// TwinCAT 3 PLC project MainPLC
// ProgramVersion: 3.1.4026.20
// libraries:
//   Tc2_Standard, * (Beckhoff Automation GmbH)
//   Tc2_System, * (Beckhoff Automation GmbH)
// project tree:
//   DUTs/ stShutterCommand.TcDUT, eShutterCommandType.TcDUT, stShutterConfig.TcDUT, eShutterStateType.TcDUT, stShutterState.TcDUT, stSwitchConfig.TcDUT, eSwitchStateType.TcDUT, stSwitchState.TcDUT
//   GVLs/ gvlSwitches.TcGVL, gvlShutters.TcGVL
//   / PlcTask.TcTTO
//   POUs/ MAIN.TcPOU
//   POUs/Shutters/ fbShutter.TcPOU, fbShutterActuator.TcPOU, fbShutterController.TcPOU
//   POUs/Switches/ fbSwitch.TcPOU
// real-time tasks:
//   TASK PlcTask: cycle T#50000us, priority 20, ADS port 350
// I/O:
//   DEVICE Device 1 (EtherCAT), AmsNetId 169.254.52.30.2.1
//     Term 4 (EK1100) [EK1100 EtherCAT Coupler (2A E-Bus)]
//       Term 5 (EL1008) [EL1008 8Ch. Dig. Input 24V, 3ms]
//       Term 6 (EL1809) [EL1809 16Ch. Dig. Input 24V, 3ms]
//       Term 7 (EL1809) [EL1809 16Ch. Dig. Input 24V, 3ms]
//       Term 8 (EL1809) [EL1809 16Ch. Dig. Input 24V, 3ms]
//       Term 9 (EL1809) [EL1809 16Ch. Dig. Input 24V, 3ms]
//       Term 10 (EL1809) [EL1809 16Ch. Dig. Input 24V, 3ms]
//       Term 11 (EL2809) [EL2809 16Ch. Dig. Output 24V, 0.5A]
//       Term 12 (EL2809) [EL2809 16Ch. Dig. Output 24V, 0.5A]
//       Term 13 (EL2809) [EL2809 16Ch. Dig. Output 24V, 0.5A]
//       Term 14 (EL2809) [EL2809 16Ch. Dig. Output 24V, 0.5A]
//       Term 15 (EL9011) [EL9011 End Terminal]
// variable links:
//   MainPLC/MainPLC Instance <-> Device 1 (EtherCAT)/Term 4 (EK1100)/Term 11 (EL2809)
//     PlcTask Outputs/gvlShutters.gvShutter1Down <-> Channel 2/Output
//     PlcTask Outputs/gvlShutters.gvShutter1Up <-> Channel 1/Output
//   MainPLC/MainPLC Instance <-> Device 1 (EtherCAT)/Term 4 (EK1100)/Term 5 (EL1008)
//     PlcTask Inputs/gvlSwitches.gvSwitchR1Down <-> Channel 2/Input
//     PlcTask Inputs/gvlSwitches.gvSwitchR1Up <-> Channel 1/Input

CONFIGURATION MainPLC
    RESOURCE PLC ON TwinCAT3
        TASK PlcTask(INTERVAL := T#50000us, PRIORITY := 20);
        PROGRAM MAIN WITH PlcTask : MAIN;
    END_RESOURCE
END_CONFIGURATION

// ---- DUTs/stShutterCommand.TcDUT
TYPE stShutterCommand :
STRUCT
    CommandType  : eShutterCommandType;	// Command type
    Position : USINT;                	// Position for MOVE_TO_POSITION command
	Angle : USINT;						// Fin Angle for MOVE_TO_POSITION command
END_STRUCT
END_TYPE

// ---- DUTs/eShutterCommandType.TcDUT
{attribute 'qualified_only'}
{attribute 'strict'}
{attribute 'to_string'}
TYPE eShutterCommandType :
(
    NONE,           // No command
    OPEN,           // Open command (move to 100%)
    CLOSE,          // Close command (move to 0%)
	STEP_OPEN,		// Open by step 10%
	STEP_CLOSE,		// Close by step 10%
    STOP,           // Stop command
    MOVE_TO_POSITION // Move to specific position
);
END_TYPE

// ---- DUTs/stShutterConfig.TcDUT
TYPE stShutterConfig :
STRUCT
    TravelTime : TIME := T#30S;			// Time for full open/close vertical movement
	AngleFullTurnTime : TIME := T#3S;			// Time for fins to make full rotation
	TravelTimeOverstep : TIME := T#500MS;		// High state output signal time allowed to be maintain after reaching full open position
END_STRUCT
END_TYPE

// ---- DUTs/eShutterStateType.TcDUT
{attribute 'qualified_only'}
{attribute 'strict'}
{attribute 'to_string'}
TYPE eShutterStateType :
(
    IDLE,            // Not moving
    MOVING_UP,       // Moving upward (opening)
    MOVING_DOWN      // Moving downward (closing)
);
END_TYPE

// ---- DUTs/stShutterState.TcDUT
TYPE stShutterState :
STRUCT
    CurrentState    : eShutterStateType;        // Current shutter state
    PreviousState   : eShutterStateType;        // Previous state
    StateChanged    : BOOL;                // State change flag
    
    CurrentPosition : USINT := 0;          // Current position [%] (0=closed, 100=open)
	CurrentAngle : USINT := 0;				// Current angle [%] (0=closed, 100=open)
    SavedPosition   : USINT := 50;         // Saved position for memory function
END_STRUCT
END_TYPE

// ---- DUTs/stSwitchConfig.TcDUT
TYPE stSwitchConfig :
STRUCT
	
    // Click timing parameters
    ShortClickMaxTime   : TIME := T#300ms;     // Max time for short click
    ShortClickDelayTime : TIME := T#300MS;     // Max time between short clicks
    LongClickMaxTime    : TIME := T#1000MS;    // Max time for long click
    
    (* Time logic:
        ShortClick < ShortClickMaxTime
        ShortClickMaxTime < LongClick < LongClickMaxTime  
        LongClickMaxTime < Hold
    *)
END_STRUCT
END_TYPE

// ---- DUTs/eSwitchStateType.TcDUT
{attribute 'qualified_only'}
{attribute 'strict'}
{attribute 'to_string'}
TYPE eSwitchStateType :
(
    IDLE,            // Idle - no action
    SHORT_CLICK,     // Short click
    LONG_CLICK,      // Long click
    HOLD_ON,         // Hold rising edge
	HOLD_OFF,		// Hold falling edge
    MULTI_CLICK      // Multiple click
);
END_TYPE

// ---- DUTs/stSwitchState.TcDUT
TYPE stSwitchState :
STRUCT
    // Logical state
    CurrentState        : eSwitchStateType;         // Current processed state
    PreviousState       : eSwitchStateType;         // Previous state
    StateChanged        : BOOL;                // State change flag
    
    // Counters
    PressCount          : USINT := 0;            // Number of clicks in sequence
    TotalPresses        : UDINT := 0;          // Total number of clicks

END_STRUCT
END_TYPE

// ---- GVLs/gvlSwitches.TcGVL
{attribute 'qualified_only'}
VAR_GLOBAL
	gvSwitchR1Up AT %I* : BOOL;
	gvSwitchR1Down AT %I* : BOOL;
END_VAR

// ---- GVLs/gvlShutters.TcGVL
{attribute 'qualified_only'}
VAR_GLOBAL
	gvShutter1Up AT %Q* : BOOL;
	gvShutter1Down AT %Q* : BOOL;
END_VAR

// ---- POUs/MAIN.TcPOU
PROGRAM MAIN
VAR
	
	PlcFirstCycle : BOOL := TRUE;

	// SWITCHES
	SwitchR1Up : fbSwitch;
	SwitchR1UpConfig : stSwitchConfig;
	SwitchR1Down : fbSwitch;
	SwitchR1DownConfig : stSwitchConfig;
	
	// SHUTTERS
	Shutter1 : fbShutter;
	Shutter1Cmd : stShutterCommand;
	Shutter1Config : stShutterConfig;
	
END_VAR


IF PlcFirstCycle THEN
	SwitchR1UpConfig.ShortClickMaxTime := T#500MS;
	SwitchR1UpConfig.ShortClickDelayTime := T#500MS;
	SwitchR1UpConfig.LongClickMaxTime := T#1500MS;
	
	SwitchR1DownConfig.ShortClickMaxTime := T#500MS;
	SwitchR1DownConfig.ShortClickDelayTime := T#500MS;
	SwitchR1DownConfig.LongClickMaxTime := T#1500MS;
	
	Shutter1Config.TravelTime := T#15S;
	Shutter1Config.AngleFullTurnTime := T#3S;
	
	PlcFirstCycle := FALSE;
END_IF


SwitchR1Up(I_Switch := gvlSwitches.gvSwitchR1Up, Config := SwitchR1UpConfig);
SwitchR1Down(I_Switch := gvlSwitches.gvSwitchR1Down, Config := SwitchR1DownConfig);

Shutter1Cmd.CommandType := eShutterCommandType.NONE;

// STOP condition - If shutter is moving, any switch R1 or R2 click will stop shutter
IF Shutter1.State.CurrentState <> eShutterStateType.IDLE AND 
	( SwitchR1Up.State.CurrentState <> eSwitchStateType.IDLE
	OR SwitchR1Down.State.CurrentState <> eSwitchStateType.IDLE) THEN
	Shutter1Cmd.CommandType := eShutterCommandType.STOP;

// OPEN condition
ELSIF SwitchR1Up.State.CurrentState = eSwitchStateType.MULTI_CLICK AND SwitchR1Up.State.PressCount = 2 THEN
	Shutter1Cmd.CommandType := eShutterCommandType.OPEN;

// Close condition
ELSIF SwitchR1Down.State.CurrentState = eSwitchStateType.MULTI_CLICK AND SwitchR1Down.State.PressCount = 2 THEN
	Shutter1Cmd.CommandType := eShutterCommandType.Close;

// STEP_OPEN condition
ELSIF SwitchR1Up.State.CurrentState = eSwitchStateType.SHORT_CLICK THEN
	Shutter1Cmd.CommandType := eShutterCommandType.STEP_OPEN;
	
// STEP_CLOSE condition
ELSIF SwitchR1Down.State.CurrentState = eSwitchStateType.SHORT_CLICK THEN
	Shutter1Cmd.CommandType := eShutterCommandType.STEP_CLOSE;
	
// MOVE_TO_POSITION condition
ELSIF SwitchR1Up.State.CurrentState = eSwitchStateType.LONG_CLICK
	OR SwitchR1Down.State.CurrentState = eSwitchStateType.LONG_CLICK THEN
	Shutter1Cmd.Position := 50;
	Shutter1Cmd.Angle := 50;
	Shutter1Cmd.CommandType := eShutterCommandType.MOVE_TO_POSITION;
END_IF

Shutter1(Command := Shutter1Cmd, Config := Shutter1Config);

gvlShutters.gvShutter1Up := Shutter1.Q_MoveUp;
gvlShutters.gvShutter1Down := Shutter1.Q_MoveDown;

END_PROGRAM

// ---- POUs/Switches/fbSwitch.TcPOU
FUNCTION_BLOCK PUBLIC fbSwitch
VAR_INPUT
	I_Switch : BOOL;							// Physical switch input
    Config : stSwitchConfig;                     // Switch configuration
END_VAR
VAR_OUTPUT
    State : stSwitchState;                   // Processed switch state
END_VAR
VAR
    // Beckhoff edge detection
    SwitchPressed : R_TRIG;                          // Rising edge detector
    SwitchReleased : F_TRIG;                          // Falling edge detector
    PressTimerQRise : R_TRIG;
	PressTimerQFall : F_TRIG;
    // Timers
    PressTimer : TON;                         // Press duration timer
    MultiClickTimer : TON;                    // Multi-click timer
    
    // Internal
    PressCount : USINT := 0;                  // Click counter
	PressTime : TIME := T#0MS;
	ClickType : eSwitchStateType := eSwitchStateType.IDLE;
END_VAR

(* 
-----------------------------
fbSwitchController:
Set State output based on Config.Input.
State persist per one PLC cycle, except IDLE, which is a default state.
Every state change sets State.StateChanged to TRUE for one PLC cycle.

SHORT_CLICK <= Config.ShortClickMaxTime
Config.ShortClickMaxTime < LONG_CLICK < Config.LongClickMaxTime
Config.LongClickMaxTime <= HOLD
MULTI_CLICK is multiple SHORT_CLICKs delayed from one another < Config.ShortClickDelayTime
State.PressCount hold amount of switch releases for MULTI_CLICK
-----------------------------
*)

ClickType := eSwitchStateType.IDLE;
State.StateChanged := FALSE;
SwitchPressed(CLK := I_Switch);
SwitchReleased(CLK := I_Switch);
PressTimerQRise(CLK := PressTimer.Q);
PressTimerQFall(CLK := PressTimer.Q);

IF SwitchPressed.Q THEN
    PressTimer(IN := TRUE, PT := Config.LongClickMaxTime);

END_IF

PressTimer();
MultiClickTimer();

IF SwitchReleased.Q THEN
	PressTime := PressTimer.ET;
	PressTimer(IN := FALSE);
	PressCount := PressCount + 1;
	MultiClickTimer(IN := FALSE);
	
	// Short click
	IF(PressTime <= Config.ShortClickMaxTime) THEN
		MultiClickTimer(IN := TRUE, PT := Config.ShortClickDelayTime);
	// Long click	
	ELSIF (PressTime < Config.LongClickMaxTime) THEN
		ClickType := eSwitchStateType.LONG_CLICK;
	// NOTE: if PressTime = Config.LongClickMaxTime, after HOLD release next state became LONG_CLICK instead of IDLE
	END_IF
END_IF

// Hold click
IF PressTimerQRise.Q THEN
    ClickType := eSwitchStateType.HOLD_ON;
END_IF

IF PressTimerQFall.Q THEN
    ClickType := eSwitchStateType.HOLD_OFF;
END_IF

IF MultiClickTimer.Q AND NOT I_Switch THEN
	IF PressCount > 1 THEN
		 ClickType := eSwitchStateType.MULTI_CLICK;
	ELSE
		ClickType := eSwitchStateType.SHORT_CLICK;
	END_IF
	MultiClickTimer(IN := FALSE);
END_IF

IF ClickType <> State.CurrentState THEN
	State.PreviousState := State.CurrentState;
	State.CurrentState := ClickType;
	State.PressCount := PressCount;
	State.StateChanged := TRUE;
	
	PressCount := 0;
END_IF

END_FUNCTION_BLOCK

// ---- POUs/Shutters/fbShutter.TcPOU
FUNCTION_BLOCK PUBLIC fbShutter
VAR_INPUT
  Command : stShutterCommand;  // Switches/HA/scheduler
  Config : stShutterConfig;
END_VAR
VAR_OUTPUT
  Q_MoveUp : BOOL;
  Q_MoveDown : BOOL;
  State : stShutterState;
END_VAR
VAR
  Ctrl : fbShutterController;
  Act : fbShutterActuator;
END_VAR

Ctrl(Command := Command, State := Act.State);
Act(MoveUp := Ctrl.MoveUp, MoveDown := Ctrl.MoveDown, Config := Config);

Q_MoveUp := Act.Q_MoveUp;
Q_MoveDown := Act.Q_MoveDown;
State := Act.State;

END_FUNCTION_BLOCK

// ---- POUs/Shutters/fbShutterController.TcPOU
FUNCTION_BLOCK PUBLIC fbShutterController
VAR_INPUT
    Command : stShutterCommand;			// Command input (one-shot or const)
	State   : stShutterState;			// Shutter state from fbShutterActuator output
END_VAR
VAR_OUTPUT
    MoveUp : BOOL;						// Signal for fbShutterActuator input
	MoveDown : BOOL;					// Signal for fbShutterActuator input
END_VAR
VAR
	CurrentCommand : stShutterCommand;
	CommandChanged : BOOL := FALSE;
	MovingToPosition : BOOL := FALSE;
	TargetPosition : USINT := 0;
	TargetAngle : USINT := 0;
END_VAR
VAR CONSTANT
	Hysteresis: USINT := 1;
	MoveStep : USINT := 10;
END_VAR

(* 
	Shutter Controller Function Block
	
	100 - fully open position/angle
	0 - fully close position/angle

*)


// Check for new command
CommandChanged := Command.CommandType <> CurrentCommand.CommandType
					OR Command.Position <> CurrentCommand.Position
					OR Command.Angle <> CurrentCommand.Angle;
					
// Handle new command
IF CommandChanged THEN
	CurrentCommand := Command;
	CASE Command.CommandType OF
		eShutterCommandType.STOP:
			MovingToPosition := FALSE;
			MoveUp := FALSE;
			MoveDown := FALSE;
			
		eShutterCommandType.OPEN:
			MovingToPosition := TRUE;
			TargetPosition := 100;
			TargetAngle := 100;
		
		eShutterCommandType.CLOSE:
			MovingToPosition := TRUE;
			TargetPosition := 0;
			TargetAngle := 0;
			
		eShutterCommandType.STEP_OPEN:
			MovingToPosition := TRUE;
			TargetPosition := State.CurrentPosition;
			// First open fins by angle step
			IF State.CurrentAngle <= 100 - MoveStep THEN
				TargetAngle := State.CurrentAngle + MoveStep;
			// If fins are fully open -> move position
			ELSE
				TargetAngle := 100;
				IF State.CurrentPosition < 100 - MoveStep THEN
					TargetPosition := State.CurrentPosition + MoveStep;
				ELSE
					TargetPosition := 100;
				END_IF
			END_IF
			//TargetPosition := State.CurrentPosition + MoveStep;
			//TargetAngle := 0;
			
		eShutterCommandType.STEP_CLOSE:
			MovingToPosition := TRUE;
			TargetPosition := State.CurrentPosition;
			// First close fins by angle step
			IF State.CurrentAngle >= 0 + MoveStep THEN
				TargetAngle := State.CurrentAngle - MoveStep;
			// If fins are fully closed -> move position
			ELSE
				TargetAngle := 0;
				IF State.CurrentPosition >= 0 + MoveStep THEN
					TargetPosition := State.CurrentPosition - MoveStep;
				ELSE
					TargetPosition := 0;
				END_IF
			END_IF
			
		eShutterCommandType.MOVE_TO_POSITION:
			MovingToPosition := TRUE;
			TargetPosition := Command.Position;
			TargetAngle := Command.Angle;
			
		eShutterCommandType.NONE:
			// No command
	END_CASE;
END_IF

IF MovingToPosition THEN	
	// Move to target vertical position first
	IF State.CurrentPosition < TargetPosition THEN
		MoveUp := TRUE;
		MoveDown := FALSE;
	ELSIF State.CurrentPosition > TargetPosition THEN
		MoveUp := FALSE;
		MoveDown := TRUE;
	ELSE
		// Then move to target angle
		IF State.CurrentAngle < TargetAngle THEN
			MoveUp := TRUE;
			MoveDown := FALSE;
		ELSIF State.CurrentAngle > TargetAngle THEN
			MoveUp := FALSE;
			MoveDown := TRUE;
		ELSE
			// Target Position and Angle achieved
			MovingToPosition := FALSE;
			MoveUp := FALSE;
			MoveDown := FALSE;
		END_IF
	END_IF
END_IF

END_FUNCTION_BLOCK

// ---- POUs/Shutters/fbShutterActuator.TcPOU
FUNCTION_BLOCK fbShutterActuator
VAR_INPUT
	MoveUp : BOOL;
	MoveDown : BOOL;
	Config : stShutterConfig;
END_VAR
VAR_OUTPUT
	Q_MoveUp : BOOL;
	Q_MoveDown : BOOL;
	State : stShutterState;
END_VAR
VAR
	OutputCheckTimer : TON;
END_VAR
VAR CONSTANT
	OutputCheckCycleTime: TIME := T#50MS;
END_VAR
VAR PERSISTENT
	CurrentPosTime: TIME := T#0S;
	CurrentAngleTime: TIME := T#0S;
END_VAR


Q_MoveUp := MoveUp;
Q_MoveDown := MoveDown;

// Both signals must not be set at the same time
IF Q_MoveUp AND Q_MoveDown THEN
	Q_MoveUp := FALSE;
	Q_MoveDown := FALSE;
END_IF

// Reset signal if shutter reached fully open position with overstep
IF Q_MoveUp AND CurrentPosTime >= Config.TravelTime + Config.TravelTimeOverstep THEN
	Q_MoveUp := FALSE;
END_IF

// Reset signal if shutter reached fully close position
IF Q_MoveDown AND CurrentPosTime <= T#0S THEN
	Q_MoveDown := FALSE;
END_IF

// Count time and accumulate when signals are set
OutputCheckTimer(IN := Q_MoveDown OR Q_MoveUp, PT := OutputCheckCycleTime);
IF OutputCheckTimer.Q THEN
	IF Q_MoveUp THEN
		// Open fins first before moving up
		IF CurrentAngleTime < Config.AngleFullTurnTime THEN
			CurrentAngleTime := CurrentAngleTime + OutputCheckCycleTime;
		ELSIF CurrentPosTime < Config.TravelTime THEN
			CurrentPosTime := CurrentPosTime + OutputCheckCycleTime;
		END_IF;
	END_IF
	
	IF Q_MoveDown THEN
		// Close fins first before moving down
		IF CurrentAngleTime > T#0S THEN
			CurrentAngleTime := CurrentAngleTime - OutputCheckCycleTime;
		ELSIF CurrentPosTime > T#0s THEN
			CurrentPosTime := CurrentPosTime - OutputCheckCycleTime;
		END_IF;
	END_IF
	
	OutputCheckTimer.IN := FALSE;  // reset
END_IF

// Update shutter position% basen on position time
State.CurrentPosition := TimeToPosition(CurrentPosTime := CurrentPosTime, TravelTime := Config.TravelTime);
State.CurrentAngle := TimeToPosition(CurrentPosTime := CurrentAngleTime, TravelTime := Config.AngleFullTurnTime);

// Update shutter current motor state
IF Q_MoveUp AND NOT Q_MoveDown THEN
	State.CurrentState := eShutterStateType.MOVING_UP;
ELSIF NOT Q_MoveUp AND Q_MoveDown THEN
	State.CurrentState := eShutterStateType.MOVING_DOWN;
ELSE
	State.CurrentState := eShutterStateType.IDLE;
END_IF

METHOD PUBLIC TimeToPosition : USINT
VAR_INPUT
	CurrentPosTime : TIME;
	TravelTime : TIME;
END_VAR
TimeToPosition := UDINT_TO_USINT(100 * TIME_TO_UDINT(CurrentPosTime) / TIME_TO_UDINT(TravelTime));
END_METHOD

END_FUNCTION_BLOCK
